(* CODESYS project Main.xml

Project tree, tasks and I/O mapping:
  visualisation Main
*)

// /Main
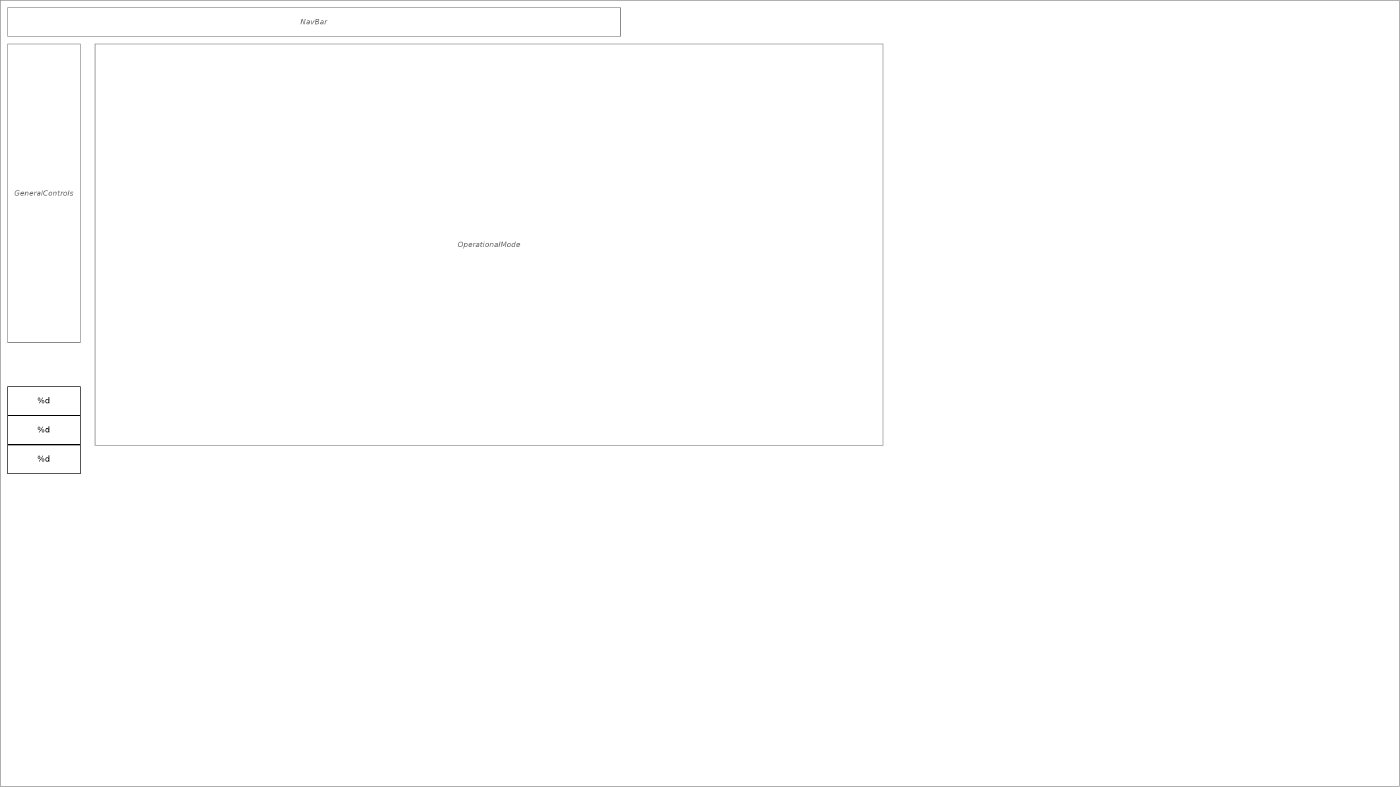
VISUALIZATION Main  // 1920x1080
    Frame (130,60 1081x551), frame switch variable: GVL_Project.fbProject._fbNavBarController.iFrame
        shows OperationalMode()
        shows SysParFeedRobot()
        shows SysParBuggy()
        shows JobManager()
        shows ManualRequest()
        shows FeedRobot()
        shows YarnStorage()
        shows SysParSafety()
        shows AxisSingle(sAxis := PRG_VisuTask_10ms._fbCreelRobotCtrl._asTitle[1], Axis := GVL_IOCContainer.fbCRAxisHw._fbAxisX)
        shows AxisSingle(sAxis := PRG_VisuTask_10ms._fbCreelRobotCtrl._asTitle[2], Axis := GVL_IOCContainer.fbCRAxisHw._fbAxisZ)
        shows AxisY()
        shows AxisSingle(sAxis := PRG_VisuTask_10ms._fbCreelRobotCtrl._asTitle[4], Axis := GVL_IOCContainer.fbCRAxisHw._fbAxisV)
        shows AxisSingle(sAxis := PRG_VisuTask_10ms._fbCreelRobotCtrl._asTitle[5], Axis := GVL_IOCContainer.fbCRAxisHw._fbAxisU)
        shows JobManager()
        shows ManualRequest()
        shows Creel()
        shows CreelRobotAxis()
        shows CreelRobotGripper()
        shows CreelRobotSplicer()
        shows CreelRobotPackageDiameter()
        shows CreelRobotCarrierDistance()
        shows CreelConveyor()
        shows Demo()
        p3621208486: PRG_VisuTask_100ms._fbCreelRobotCtrl._asTitle[2]
        p182062315: GVL_IOCContainer.fbCreelRobot._fbRobotAxis._fbAxisZ
    Rectangle (10,530 100x40), "%d", text variable: PRG_PlcTask_10ms._iHeartBeat
    Rectangle (10,570 100x40), "%d", text variable: PRG_PlcTask_50ms._iHeartBeat
    Rectangle (10,610 100x40), "%d", text variable: PRG_VisuTask_100ms._iHeartBeat
    Frame (10,10 841x40)
        shows NavBar()
    Frame (10,60 100x410)
        shows GeneralControls()
END_VISUALIZATION
